Fanuc KAREL source: KA00069.KL

PROGRAM KA00069
%NOLOCKGROUP
VAR
  SRC: XYZWPR
  DST: VECTOR
BEGIN
  SRC.X = 1.0
  DST = SRC
END KA00069
